FUNCTION_BLOCK fbStepToTarget
VAR_INPUT
    TargetVal : USINT;
    StepVal : USINT;
    CycleTime : TIME;
END_VAR
VAR_IN_OUT
    Value : USINT;
END_VAR
VAR_OUTPUT
    Reached : BOOL;
END_VAR
VAR
    StepTimer : TON;
END_VAR

(*
	Increment/Decrement Value by StepVal every CycleTime until it reaches TargetVal.
	After reaching TargetVal set Reached for one cycle
*)

Reached := FALSE;

IF StepVal <= 0.0 THEN
    RETURN;
END_IF

StepTimer(IN := TRUE, PT := CycleTime);

IF Value < TargetVal THEN
    IF StepTimer.Q THEN
        Value := Value + StepVal;
        IF Value >= TargetVal THEN
            Value := TargetVal;
            Reached := TRUE;
        END_IF
        StepTimer(IN := FALSE);
    END_IF

ELSIF Value > TargetVal THEN
    IF StepTimer.Q THEN
        Value := Value - StepVal;
        IF Value <= TargetVal THEN
            Value := TargetVal;
            Reached := TRUE;
        END_IF
        StepTimer(IN := FALSE);
    END_IF
END_IF

END_FUNCTION_BLOCK

(* stored: Version 1.1.0.1
   POU fbStepToTarget: Id {139c758d-a096-42f2-b819-2ba7838a396f}, SpecialFunc None *)
